(* IEC 61131-3 sources: avi-aoi-management/scripts/ai-eval/ngau-nhien/lib/st-scl/mau-scl/st-ud8-pi-chong-bao-hoa/src, 2 files *)

(* ---- KepGioiHan.st ---- *)
FUNCTION "KepGioiHan" : Real
{ S7_Optimized_Access := 'TRUE' }
VERSION : 0.1
   VAR_INPUT
      X : Real;
      LO : Real;
      HI : Real;
   END_VAR

BEGIN
   IF #X < #LO THEN
      #KepGioiHan := #LO;
   ELSIF #X > #HI THEN
      #KepGioiHan := #HI;
   ELSE
      #KepGioiHan := #X;
   END_IF;
END_FUNCTION

(* ---- BoPI.st ---- *)
FUNCTION_BLOCK "BoPI"
{ S7_Optimized_Access := 'TRUE' }
VERSION : 0.1
   VAR_INPUT
      SP : Real;
      PV : Real;
      KP : Real;
      TI : Real;
      TS : Time;
      U_MIN : Real;
      U_MAX : Real;
      MAN : Bool;
      U_TAY : Real;
   END_VAR

   VAR_OUTPUT
      U : Real;
      I_TP : Real;
      BAO_HOA_CAO : Bool;
      BAO_HOA_THAP : Bool;
   END_VAR

   VAR
      tTruoc : Time;
      daTinh : Bool;
   END_VAR

   VAR_TEMP
      e : Real;
      uTho : Real;
      tsGiay : Real;
   END_VAR

BEGIN
   #e := #SP - #PV;
   IF #MAN THEN
      // Tay: U theo U_TAY, tích phân bám để chuyển về tự động không giật
      #U := "KepGioiHan"(X := #U_TAY, LO := #U_MIN, HI := #U_MAX);
      #I_TP := #U - #KP * #e;
      #BAO_HOA_CAO := FALSE;
      #BAO_HOA_THAP := FALSE;
      #tTruoc := "G_NOW";
      #daTinh := TRUE;
   ELSIF NOT #daTinh OR ("G_NOW" - #tTruoc >= #TS) THEN
      #tTruoc := "G_NOW";
      #daTinh := TRUE;
      #tsGiay := LINT_TO_REAL(TIME_TO_LINT(#TS)) / 1.0E9;
      #uTho := #KP * #e + #I_TP;
      #BAO_HOA_CAO := #uTho > #U_MAX;
      #BAO_HOA_THAP := #uTho < #U_MIN;
      // Chống bão hoà: không tích phân thêm theo chiều đang bão hoà
      IF NOT ((#BAO_HOA_CAO AND #e > 0.0) OR (#BAO_HOA_THAP AND #e < 0.0)) THEN
         #I_TP := #I_TP + #KP * #tsGiay / #TI * #e;
      END_IF;
      #U := "KepGioiHan"(X := #uTho, LO := #U_MIN, HI := #U_MAX);
   END_IF;
END_FUNCTION_BLOCK
